TYPE ST_VC_InspectionResult :
STRUCT
    Pass          : BOOL;
    ErrorCode     : DINT;
    MeasuredCount : UINT;
    Measured      : ARRAY[0..15] OF REAL;
END_STRUCT
END_TYPE

(* stored: Version 1.1.0.1, ProductVersion 3.1.4026.21
   DUT ST_VC_InspectionResult: Id {ebad5a86-5b59-4a03-b820-3a2abd2c5375} *)
